FUNCTION_BLOCK F (* Negative C5: two positions that only toggle and run the same algorithm *)
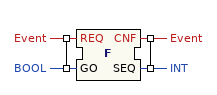
  EVENT_INPUT
    REQ WITH GO;
  END_EVENT
  EVENT_OUTPUT
    CNF WITH SEQ;
  END_EVENT
  VAR_INPUT
    GO : BOOL;
  END_VAR
  VAR_OUTPUT
    SEQ : INT;
  END_VAR
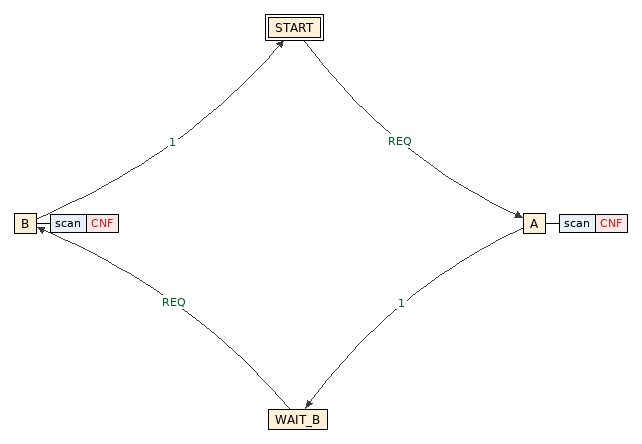
  EC_STATES
    START;
    A : scan -> CNF;
    WAIT_B;
    B : scan -> CNF;
  END_STATES
  EC_TRANSITIONS
    START TO A := REQ;
    A TO WAIT_B := 1;
    WAIT_B TO B := REQ;
    B TO START := 1;
  END_TRANSITIONS
  ALGORITHM scan IN ST:
IF GO THEN
  SEQ := 1;
ELSE
  SEQ := 0;
END_IF;
  END_ALGORITHM
END_FUNCTION_BLOCK
